    - item type 7 BRTIRUS1510A : 21 | -6861
    - item type 7 BRTIRUS1510A : 21 | -6862
    - item type 7 BRTIRUS1510A : 21 | -6863
    - item type 7 BRTIRUS1510A : 21 | -6864
    - item type 7 BRTIRUS1510A : 21 | -6865
    - item type 7 BRTIRUS1510A : 21 | -6866
    - item type 7 BRTIRUS1510A : 21 | -6867
    - item type 7 BRTIRUS1510A : 21 | -6868
    - item type 7 BRTIRUS1510A : 21 | -6869
    - item type 7 BRTIRUS1510A : 21 | -6870
    - item type 7 BRTIRUS1510A : 21 | -6871
    - item type 7 BRTIRUS1510A : 21 | -6872
    - item type 7 BRTIRUS1510A : 21 | -6873
    - item type 7 BRTIRUS1510A : 21 | -6874
    - item type 7 BRTIRUS1510A : 21 | -6875
    - item type 7 BRTIRUS1510A : 21 | -6876
    - item type 7 BRTIRUS1510A : 21 | -6877
    - item type 7 BRTIRUS1510A : 21 | -6878
    - item type 7 BRTIRUS1510A : 21 | -6879
    - item type 7 BRTIRUS1510A : 21 | -6880
    - item type 7 BRTIRUS1510A : 21 | -6881
    - item type 7 BRTIRUS1510A : 21 | -6882
    - item type 7 BRTIRUS1510A : 21 | -6883
    - item type 7 BRTIRUS1510A : 21 | -6884
    - item type 7 BRTIRUS1510A : 21 | -6885
    - item type 7 BRTIRUS1510A : 21 | -6886
    - item type 7 BRTIRUS1510A : 21 | -6887
    - item type 7 BRTIRUS1510A : 21 | -6888
    - item type 7 BRTIRUS1510A : 21 | -6889
    - item type 7 BRTIRUS1510A : 21 | -6890
    - item type 7 BRTIRUS1510A : 21 | -6891
    - item type 7 BRTIRUS1510A : 21 | -6892
    - item type 7 BRTIRUS1510A : 21 | -6893
    - item type 7 BRTIRUS1510A : 21 | -6894
    - item type 7 BRTIRUS1510A : 21 | -6895
    - item type 7 BRTIRUS1510A : 21 | -6896
    - item type 7 BRTIRUS1510A : 21 | -6897
    - item type 7 BRTIRUS1510A : 21 | -6898
    - item type 7 BRTIRUS1510A : 21 | -6899
    - item type 7 BRTIRUS1510A : 21 | -6900
    - item type 7 BRTIRUS1510A : 21 | -6901
    - item type 7 BRTIRUS1510A : 21 | -6902
    - item type 7 BRTIRUS1510A : 21 | -6903
    - item type 7 BRTIRUS1510A : 21 | -6904
    - item type 7 BRTIRUS1510A : 21 | -6905
    - item type 7 BRTIRUS1510A : 21 | -6906
    - item type 7 BRTIRUS1510A : 21 | -6907
    - item type 7 BRTIRUS1510A : 21 | -6908
    - item type 7 BRTIRUS1510A : 21 | -6909
    - item type 7 BRTIRUS1510A : 21 | -6910
    - item type 7 BRTIRUS1510A : 21 | -6911
    - item type 7 BRTIRUS1510A : 21 | -6912
    - item type 7 BRTIRUS1510A : 21 | -6913
    - item type 7 BRTIRUS1510A : 21 | -6914
    - item type 7 BRTIRUS1510A : 21 | -6915
    - item type 7 BRTIRUS1510A : 21 | -6916
    - item type 7 BRTIRUS1510A : 21 | -6917
    - item type 7 BRTIRUS1510A : 21 | -6918
    - item type 7 BRTIRUS1510A : 21 | -6919
    - item type 7 BRTIRUS1510A : 21 | -6920
    - item type 7 BRTIRUS1510A : 21 | -6921
    - item type 7 BRTIRUS1510A : 21 | -6922
    - item type 7 BRTIRUS1510A : 21 | -6923
    - item type 7 BRTIRUS1510A : 21 | -6924
    - item type 7 BRTIRUS1510A : 21 | -6925
    - item type 7 BRTIRUS1510A : 21 | -6926
    - item type 7 BRTIRUS1510A : 21 | -6927
    - item type 7 BRTIRUS1510A : 21 | -6928
    - item type 7 BRTIRUS1510A : 21 | -6929
    - item type 7 BRTIRUS1510A : 21 | -6930
    - item type 7 BRTIRUS1510A : 21 | -6931
    - item type 7 BRTIRUS1510A : 21 | -6932
    - item type 7 BRTIRUS1510A : 21 | -6933
    - item type 7 BRTIRUS1510A : 21 | -6934
    - item type 7 BRTIRUS1510A : 21 | -6935
    - item type 7 BRTIRUS1510A : 21 | -6936
    - item type 7 BRTIRUS1510A : 21 | -6937
    - item type 7 BRTIRUS1510A : 21 | -6938
    - item type 7 BRTIRUS1510A : 21 | -6939
    - item type 7 BRTIRUS1510A : 21 | -6940
    - item type 7 BRTIRUS1510A : 21 | -6941
    - item type 7 BRTIRUS1510A : 21 | -6942
    - item type 7 BRTIRUS1510A : 21 | -6943
    - item type 7 BRTIRUS1510A : 21 | -6944
    - item type 7 BRTIRUS1510A : 21 | -6945
    - item type 7 BRTIRUS1510A : 21 | -6946
    - item type 7 BRTIRUS1510A : 21 | -6947
    - item type 7 BRTIRUS1510A : 21 | -6948
    - item type 7 BRTIRUS1510A : 21 | -6949
    - item type 7 BRTIRUS1510A : 21 | -6950
    - item type 7 BRTIRUS1510A : 21 | -6951
    - item type 7 BRTIRUS1510A : 21 | -6952
    - item type 7 BRTIRUS1510A : 21 | -6953
    - item type 7 BRTIRUS1510A : 21 | -6954
    - item type 7 BRTIRUS1510A : 21 | -6955
    - item type 7 BRTIRUS1510A : 21 | -6956
    - item type 7 BRTIRUS1510A : 21 | -6957
    - item type 7 BRTIRUS1510A : 21 | -6958
    - item type 7 BRTIRUS1510A : 21 | -6959
    - item type 7 BRTIRUS1510A : 21 | -6960
    - item type 7 BRTIRUS1510A : 21 | -6961
    - item type 7 BRTIRUS1510A : 21 | -6962
    - item type 7 BRTIRUS1510A : 21 | -6963
    - item type 7 BRTIRUS1510A : 21 | -6964
    - item type 7 BRTIRUS1510A : 21 | -6965
    - item type 7 BRTIRUS1510A : 21 | -6966
    - item type 7 BRTIRUS1510A : 21 | -6967
    - item type 7 BRTIRUS1510A : 21 | -6968
    - item type 7 BRTIRUS1510A : 21 | -6969
    - item type 7 BRTIRUS1510A : 21 | -6970
    - item type 7 BRTIRUS1510A : 21 | -6971
    - item type 7 BRTIRUS1510A : 21 | -6972
    - item type 7 BRTIRUS1510A : 21 | -6973
    - item type 7 BRTIRUS1510A : 21 | -6974
    - item type 7 BRTIRUS1510A : 21 | -6975
    - item type 7 BRTIRUS1510A : 21 | -6976
    - item type 7 BRTIRUS1510A : 21 | -6977
    - item type 7 BRTIRUS1510A : 21 | -6978
    - item type 7 BRTIRUS1510A : 21 | -6979
    - item type 7 BRTIRUS1510A : 21 | -6980
    - item type 7 BRTIRUS1510A : 21 | -6981
    - item type 7 BRTIRUS1510A : 21 | -6982
    - item type 7 BRTIRUS1510A : 21 | -6983
    - item type 7 BRTIRUS1510A : 21 | -6984
    - item type 7 BRTIRUS1510A : 21 | -6985
    - item type 7 BRTIRUS1510A : 21 | -6986
    - item type 7 BRTIRUS1510A : 21 | -6987
    - item type 7 BRTIRUS1510A : 21 | -6988
    - item type 7 BRTIRUS1510A : 21 | -6989
    - item type 7 BRTIRUS1510A : 21 | -6990
    - item type 7 BRTIRUS1510A : 21 | -6991
    - item type 7 BRTIRUS1510A : 21 | -6992
    - item type 7 BRTIRUS1510A : 21 | -6993
    - item type 7 BRTIRUS1510A : 21 | -6994
    - item type 7 BRTIRUS1510A : 21 | -6995
    - item type 7 BRTIRUS1510A : 21 | -6996
    - item type 7 BRTIRUS1510A : 21 | -6997
    - item type 7 BRTIRUS1510A : 21 | -6998
    - item type 7 BRTIRUS1510A : 21 | -6999
    - item type 7 BRTIRUS1510A : 21 | -7000
    - item type 7 BRTIRUS1510A : 21 | -7001
    - item type 7 BRTIRUS1510A : 21 | -7002
    - item type 7 BRTIRUS1510A : 21 | -7003
    - item type 7 BRTIRUS1510A : 21 | -7004
    - item type 7 BRTIRUS1510A : 21 | -7005
    - item type 7 BRTIRUS1510A : 21 | -7006
    - item type 7 BRTIRUS1510A : 21 | -7007
    - item type 7 BRTIRUS1510A : 21 | -7008
    - item type 7 BRTIRUS1510A : 21 | -7009
    - item type 7 BRTIRUS1510A : 21 | -7010
    - item type 7 BRTIRUS1510A : 21 | -7011
    - item type 7 BRTIRUS1510A : 21 | -7012
    - item type 7 BRTIRUS1510A : 21 | -7013
    - item type 7 BRTIRUS1510A : 21 | -7014
    - item type 7 BRTIRUS1510A : 21 | -7015
    - item type 7 BRTIRUS1510A : 21 | -7016
    - item type 7 BRTIRUS1510A : 21 | -7017
    - item type 7 BRTIRUS1510A : 21 | -7018
    - item type 7 BRTIRUS1510A : 21 | -7019
    - item type 7 BRTIRUS1510A : 21 | -7020
    - item type 7 BRTIRUS1510A : 21 | -7021
    - item type 7 BRTIRUS1510A : 21 | -7022
    - item type 7 BRTIRUS1510A : 21 | -7023
    - item type 7 BRTIRUS1510A : 21 | -7024
    - item type 7 BRTIRUS1510A : 21 | -7025
    - item type 7 BRTIRUS1510A : 21 | -7026
    - item type 7 BRTIRUS1510A : 21 | -7027
    - item type 7 BRTIRUS1510A : 21 | -7028
    - item type 7 BRTIRUS1510A : 21 | -7029
    - item type 7 BRTIRUS1510A : 21 | -7030
    - item type 7 BRTIRUS1510A : 21 | -7031
    - item type 7 BRTIRUS1510A : 21 | -7032
    - item type 7 BRTIRUS1510A : 21 | -7033
    - item type 7 BRTIRUS1510A : 21 | -7034
    - item type 7 BRTIRUS1510A : 21 | -7035
    - item type 7 BRTIRUS1510A : 21 | -7036
    - item type 7 BRTIRUS1510A : 21 | -7037
    - item type 7 BRTIRUS1510A : 21 | -7038
    - item type 7 BRTIRUS1510A : 21 | -7039
    - item type 7 BRTIRUS1510A : 21 | -7040
    - item type 7 BRTIRUS1510A : 21 | -7041
    - item type 7 BRTIRUS1510A : 21 | -7042
    - item type 7 BRTIRUS1510A : 21 | -7043
    - item type 7 BRTIRUS1510A : 21 | -7044
    - item type 7 BRTIRUS1510A : 21 | -7045
    - item type 7 BRTIRUS1510A : 21 | -7046
    - item type 7 BRTIRUS1510A : 21 | -7047
    - item type 7 BRTIRUS1510A : 21 | -7048
  - object BRT_Base at (0, 0, 0) mm, size 594 x 395 x 235 mm
  - object BRT_Link1 at (0, 0, 0) mm, size 483.3 x 356.2 x 433.6 mm
  - object BRT_Link2 at (0, 0, 0) mm, size 261.9 x 165.2 x 873 mm
  - object BRT_Link3 at (0, 0, 0) mm, size 320.1 x 281.6 x 342 mm
  - object BRT_Link4 at (0, 0, 0) mm, size 558.6 x 157.8 x 191.9 mm
  - object BRT_Link5 at (0, 0, 0) mm, size 153.5 x 104.8 x 120.9 mm
  - object BRT_Link6 at (0, 0, 0) mm, size 23.9 x 58.3 x 62.9 mm
  - frame BORUNTE_BRTIRUS1510A Base at (0, 0, -175) mm
    - robot BORUNTE_BRTIRUS1510A: 6 axes, payload 10 kg, weight 152 kg
        modified DH rows (alpha deg, a mm, theta deg, d mm): 0, 0, 0, 488; -90, 170, -90, 0; 0, 650, 0, 0; -90, 162, 0, 634.4; 90, 0, 0, 0; -90, 0, 0, 117
        joint limits [-165, -95, -85, -180, -115, -360] to [165, 70, 75, 180, 115, 360]; home [0, 0, 0, 0, 0, 0]; saved at [0, -1.219, 5.316, 0, 0.15, 0]
      - tool tool du an, TCP at (-221, 0, 59.5) mm, rotated rx 0 ry -90 rz 0 deg, size 140 x 350 x 102 mm, geometry from tool du an.STEP
